{attribute 'qualified_only'}
VAR_GLOBAL
    stLivingRoomCeilingRelayId : ST_DeviceId := (sId := 201, sName := 'Ceiling Relay', sRoom := 'Living Room');
    stLivingRoomWallRelayId    : ST_DeviceId := (sId := 202, sName := 'Wall Relay', sRoom := 'Living Room');
    stLivingRoomAmbientRelayId : ST_DeviceId := (sId := 203, sName := 'Ambient Relay', sRoom := 'Living Room');

    fbLivingRoomCeilingRelay : FB_RelayMonostable;
    fbLivingRoomWallRelay    : FB_RelayMonostable;
    fbLivingRoomAmbientRelay : FB_RelayMonostable;

    stLivingRoomCeilingId : ST_DeviceId := (sId := 301, sName := 'Ceiling Light', sRoom := 'Living Room');
    stLivingRoomWallId    : ST_DeviceId := (sId := 302, sName := 'Wall Light', sRoom := 'Living Room');
    stLivingRoomAmbientId : ST_DeviceId := (sId := 303, sName := 'Ambient Light', sRoom := 'Living Room');

    fbLivingRoomCeiling : FB_Light;
    fbLivingRoomWall    : FB_Light;
    fbLivingRoomAmbient : FB_Light;
END_VAR

(* stored: Version 1.1.0.1, ProductVersion 3.1.4026.20
   GVL GVL_Lights: Id {A8100002-3B71-4C96-8F25-7A1B2C3D4001} *)
